(* IEC 61131-3 sources: codesys-ai-industrial-robot-control/plc/src/Process/FB_SortingCell, 2 files *)

(* ---- AlarmState.st ---- *)
// State of one alarm (for the HMI view).
METHOD AlarmState : ST_Alarm
VAR_INPUT
    eId : E_AlarmId;
END_VAR

AlarmState := fbAlarms.GetAlarm(eId);

(* ---- PlacedCount.st ---- *)
// Parts placed in all bins since the last reset of the counters.
METHOD PlacedCount : UINT
VAR
    eBin : E_Bin;
END_VAR

PlacedCount := 0;
FOR eBin := E_Bin.TypeA TO E_Bin.Quarantine DO
    PlacedCount := PlacedCount + aBins[eBin].uiCount;
END_FOR
